(* Schneider Machine Expert - Basic project timer_options_behavior, file version 3.0.0.0 *)
(* ProjectInformations: Name=New project *)

HARDWARE
  Cpu 0: TM200CE40T
  EthernetConfiguration: NetworkName=M200, IpAllocationMode=FixedAddress, IpAddress=0.0.0.0, SubnetMask=0.0.0.0
  SerialLineConfiguration: Baud=Baud19200, Parity=ParityEven, DataBits=DataBits8, StopBits=StopBits1, PhysicalMedium=PhysicalMediumRs485, TransmissionMode=TransmissionModeModbusRtu, SlaveId=1, Addressing=SlaveAddressing
  MastTask: UsePeriodScanMode=false, PeriodScan=100
  FastTask: Period=255
  CpuBehavior: StartingMode=StartAsPreviousState, AutoSaveRamOnEeprom=true, WatchdogPeriod=250

SYMBOLS  (address, symbol, comment, settings)
  %M500     constant_false_500
  %M501     compiler_reused_M501_501
  %M502     compiler_reused_M502_502
  %M503     compiler_reused_M503_503
  %M504     compiler_reused_M504_504
  %M505     compiler_reused_M505_505
  %M506     compiler_reused_M506_506
  %M507     compiler_reused_M507_507
  %M508     compiler_reused_M508_508
  %M509     compiler_reused_M509_509
  %M510     output_5_image_510
  %M511     input_1_snapshot_511
  %M512     output_6_image_512
  %M513     input_0_snapshot_513
  %M514     output_7_image_514
  %M515     output_8_image_515
  %M516     output_9_image_516
  %M517     output_10_image_517
  %M518     output_11_image_518
  %M519     output_12_image_519
  %M520     output_13_image_520
  %M521     output_14_image_521
  %S13      SB_FIRSTRUN  "Indicates the first controller cycle in RUN mode"
  %MW4000   compiler_reused_MW4000_MW4000
  %TM0        [Preset=20, Base=OneSecond, IsRetentive=true]
  %TM1        [Type=TOF, Preset=20, Base=OneSecond, IsRetentive=true]
  %TM2        [Preset=20, Base=OneSecond, IsDynamicPreset=true]

POU Generated C++ - EXPERIMENTAL
  (* SectionNumber=1 *)

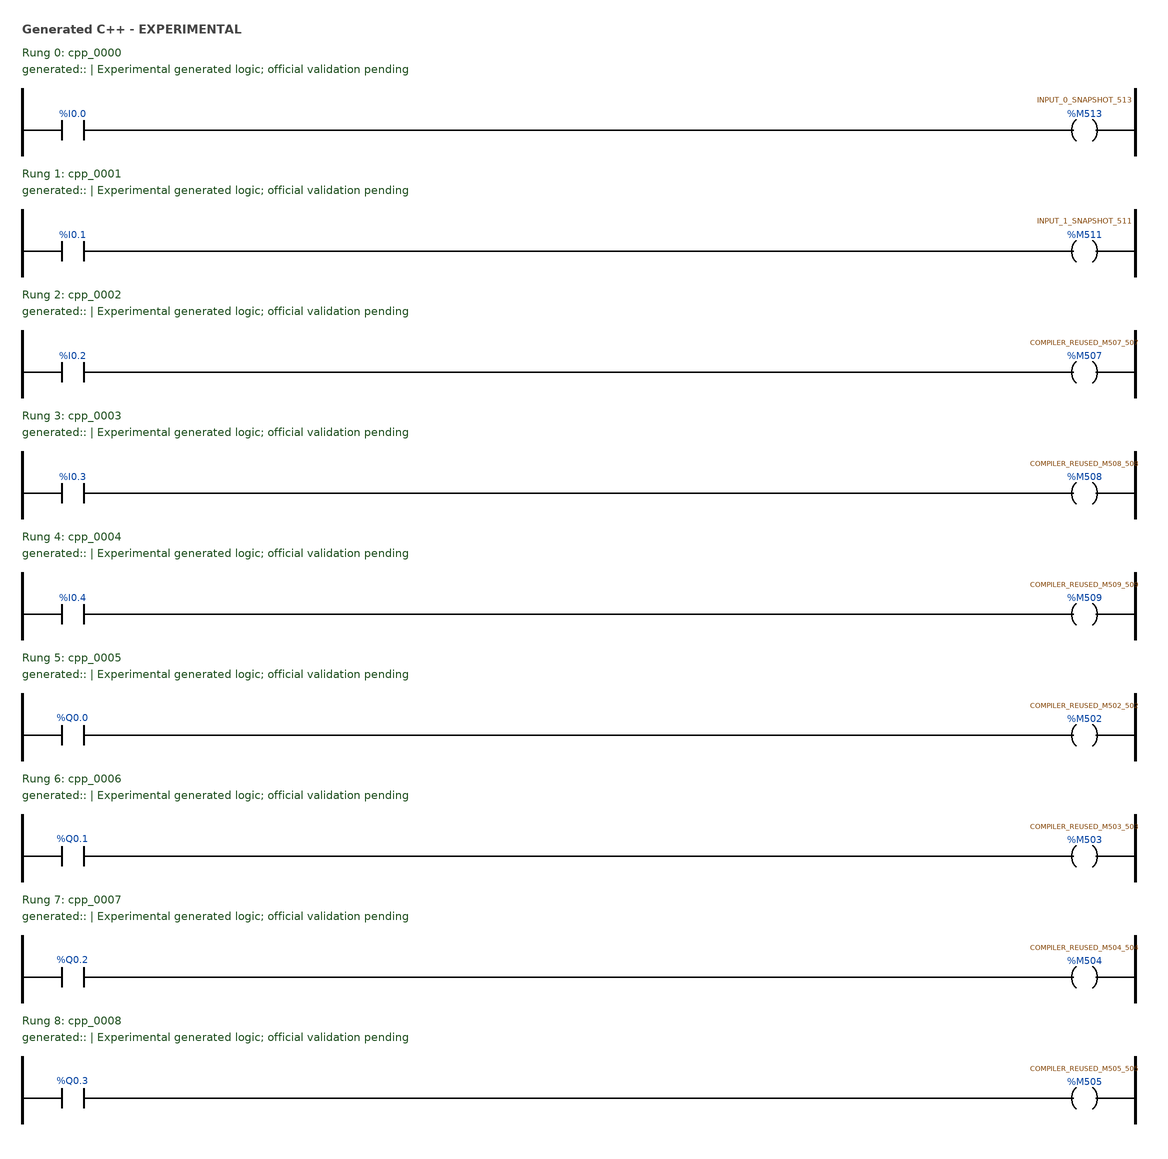

// Rung 0: cpp_0000
// generated:: | Experimental generated logic; official validation pending
  LD %I0.0
  ST %M513                (* input_0_snapshot_513 *)
  // as ST:
  //   input_0_snapshot_513 := %I0.0;

// Rung 1: cpp_0001
// generated:: | Experimental generated logic; official validation pending
  LD %I0.1
  ST %M511                (* input_1_snapshot_511 *)
  // as ST:
  //   input_1_snapshot_511 := %I0.1;

// Rung 2: cpp_0002
// generated:: | Experimental generated logic; official validation pending
  LD %I0.2
  ST %M507                (* compiler_reused_M507_507 *)
  // as ST:
  //   compiler_reused_M507_507 := %I0.2;

// Rung 3: cpp_0003
// generated:: | Experimental generated logic; official validation pending
  LD %I0.3
  ST %M508                (* compiler_reused_M508_508 *)
  // as ST:
  //   compiler_reused_M508_508 := %I0.3;

// Rung 4: cpp_0004
// generated:: | Experimental generated logic; official validation pending
  LD %I0.4
  ST %M509                (* compiler_reused_M509_509 *)
  // as ST:
  //   compiler_reused_M509_509 := %I0.4;

// Rung 5: cpp_0005
// generated:: | Experimental generated logic; official validation pending
  LD %Q0.0
  ST %M502                (* compiler_reused_M502_502 *)
  // as ST:
  //   compiler_reused_M502_502 := %Q0.0;

// Rung 6: cpp_0006
// generated:: | Experimental generated logic; official validation pending
  LD %Q0.1
  ST %M503                (* compiler_reused_M503_503 *)
  // as ST:
  //   compiler_reused_M503_503 := %Q0.1;

// Rung 7: cpp_0007
// generated:: | Experimental generated logic; official validation pending
  LD %Q0.2
  ST %M504                (* compiler_reused_M504_504 *)
  // as ST:
  //   compiler_reused_M504_504 := %Q0.2;

// Rung 8: cpp_0008
// generated:: | Experimental generated logic; official validation pending
  LD %Q0.3
  ST %M505                (* compiler_reused_M505_505 *)
  // as ST:
  //   compiler_reused_M505_505 := %Q0.3;

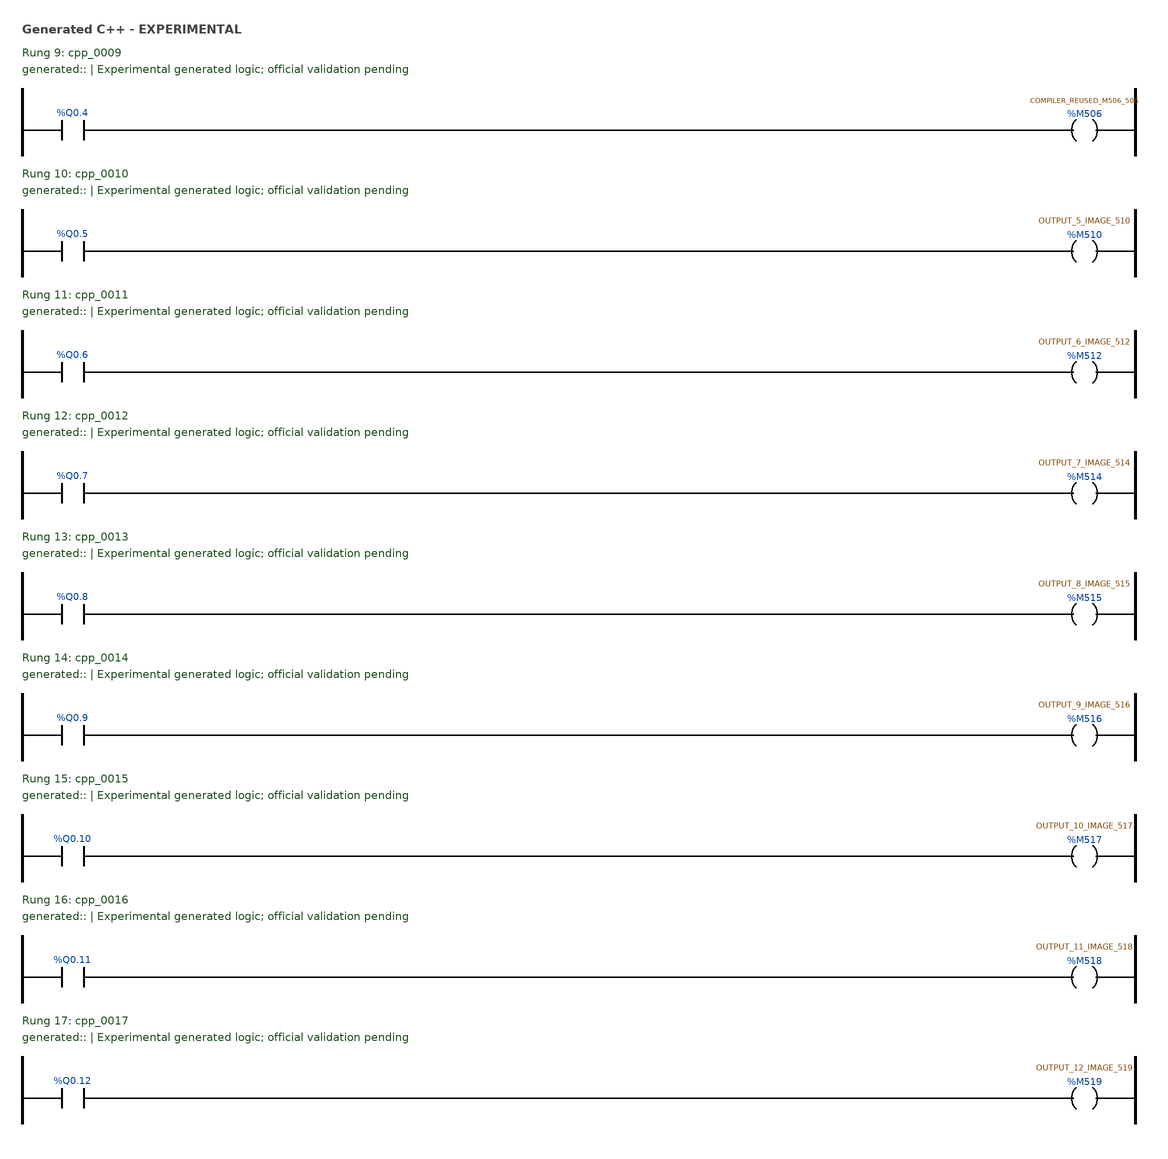

// Rung 9: cpp_0009
// generated:: | Experimental generated logic; official validation pending
  LD %Q0.4
  ST %M506                (* compiler_reused_M506_506 *)
  // as ST:
  //   compiler_reused_M506_506 := %Q0.4;

// Rung 10: cpp_0010
// generated:: | Experimental generated logic; official validation pending
  LD %Q0.5
  ST %M510                (* output_5_image_510 *)
  // as ST:
  //   output_5_image_510 := %Q0.5;

// Rung 11: cpp_0011
// generated:: | Experimental generated logic; official validation pending
  LD %Q0.6
  ST %M512                (* output_6_image_512 *)
  // as ST:
  //   output_6_image_512 := %Q0.6;

// Rung 12: cpp_0012
// generated:: | Experimental generated logic; official validation pending
  LD %Q0.7
  ST %M514                (* output_7_image_514 *)
  // as ST:
  //   output_7_image_514 := %Q0.7;

// Rung 13: cpp_0013
// generated:: | Experimental generated logic; official validation pending
  LD %Q0.8
  ST %M515                (* output_8_image_515 *)
  // as ST:
  //   output_8_image_515 := %Q0.8;

// Rung 14: cpp_0014
// generated:: | Experimental generated logic; official validation pending
  LD %Q0.9
  ST %M516                (* output_9_image_516 *)
  // as ST:
  //   output_9_image_516 := %Q0.9;

// Rung 15: cpp_0015
// generated:: | Experimental generated logic; official validation pending
  LD %Q0.10
  ST %M517                (* output_10_image_517 *)
  // as ST:
  //   output_10_image_517 := %Q0.10;

// Rung 16: cpp_0016
// generated:: | Experimental generated logic; official validation pending
  LD %Q0.11
  ST %M518                (* output_11_image_518 *)
  // as ST:
  //   output_11_image_518 := %Q0.11;

// Rung 17: cpp_0017
// generated:: | Experimental generated logic; official validation pending
  LD %Q0.12
  ST %M519                (* output_12_image_519 *)
  // as ST:
  //   output_12_image_519 := %Q0.12;

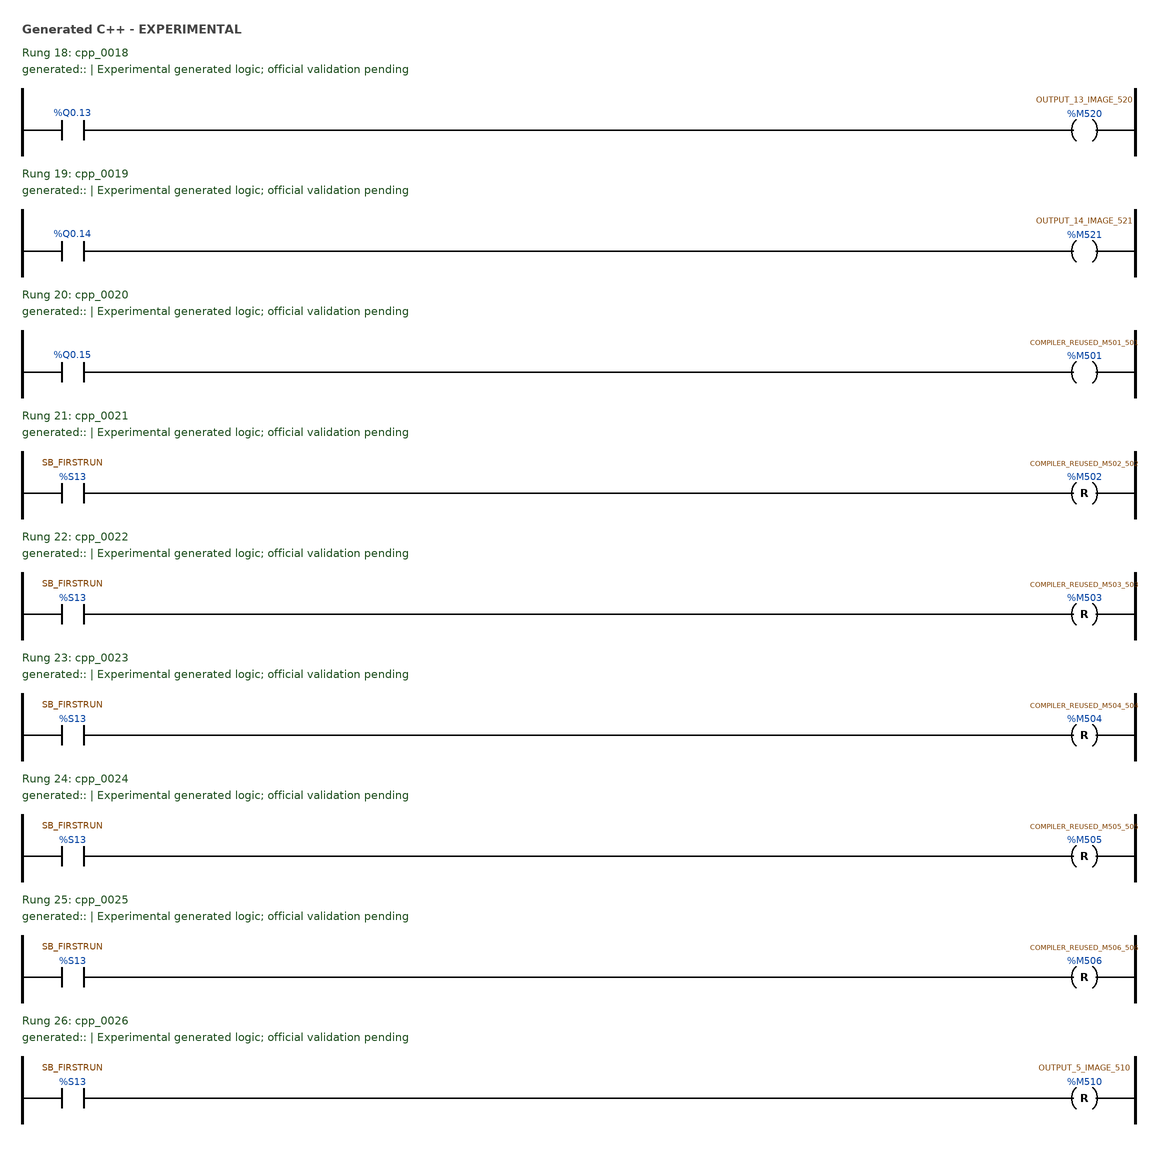

// Rung 18: cpp_0018
// generated:: | Experimental generated logic; official validation pending
  LD %Q0.13
  ST %M520                (* output_13_image_520 *)
  // as ST:
  //   output_13_image_520 := %Q0.13;

// Rung 19: cpp_0019
// generated:: | Experimental generated logic; official validation pending
  LD %Q0.14
  ST %M521                (* output_14_image_521 *)
  // as ST:
  //   output_14_image_521 := %Q0.14;

// Rung 20: cpp_0020
// generated:: | Experimental generated logic; official validation pending
  LD %Q0.15
  ST %M501                (* compiler_reused_M501_501 *)
  // as ST:
  //   compiler_reused_M501_501 := %Q0.15;

// Rung 21: cpp_0021
// generated:: | Experimental generated logic; official validation pending
  LD %S13                 (* SB_FIRSTRUN *)
  R %M502                 (* compiler_reused_M502_502 *)
  // as ST:
  //   IF SB_FIRSTRUN THEN compiler_reused_M502_502 := FALSE; END_IF;

// Rung 22: cpp_0022
// generated:: | Experimental generated logic; official validation pending
  LD %S13                 (* SB_FIRSTRUN *)
  R %M503                 (* compiler_reused_M503_503 *)
  // as ST:
  //   IF SB_FIRSTRUN THEN compiler_reused_M503_503 := FALSE; END_IF;

// Rung 23: cpp_0023
// generated:: | Experimental generated logic; official validation pending
  LD %S13                 (* SB_FIRSTRUN *)
  R %M504                 (* compiler_reused_M504_504 *)
  // as ST:
  //   IF SB_FIRSTRUN THEN compiler_reused_M504_504 := FALSE; END_IF;

// Rung 24: cpp_0024
// generated:: | Experimental generated logic; official validation pending
  LD %S13                 (* SB_FIRSTRUN *)
  R %M505                 (* compiler_reused_M505_505 *)
  // as ST:
  //   IF SB_FIRSTRUN THEN compiler_reused_M505_505 := FALSE; END_IF;

// Rung 25: cpp_0025
// generated:: | Experimental generated logic; official validation pending
  LD %S13                 (* SB_FIRSTRUN *)
  R %M506                 (* compiler_reused_M506_506 *)
  // as ST:
  //   IF SB_FIRSTRUN THEN compiler_reused_M506_506 := FALSE; END_IF;

// Rung 26: cpp_0026
// generated:: | Experimental generated logic; official validation pending
  LD %S13                 (* SB_FIRSTRUN *)
  R %M510                 (* output_5_image_510 *)
  // as ST:
  //   IF SB_FIRSTRUN THEN output_5_image_510 := FALSE; END_IF;

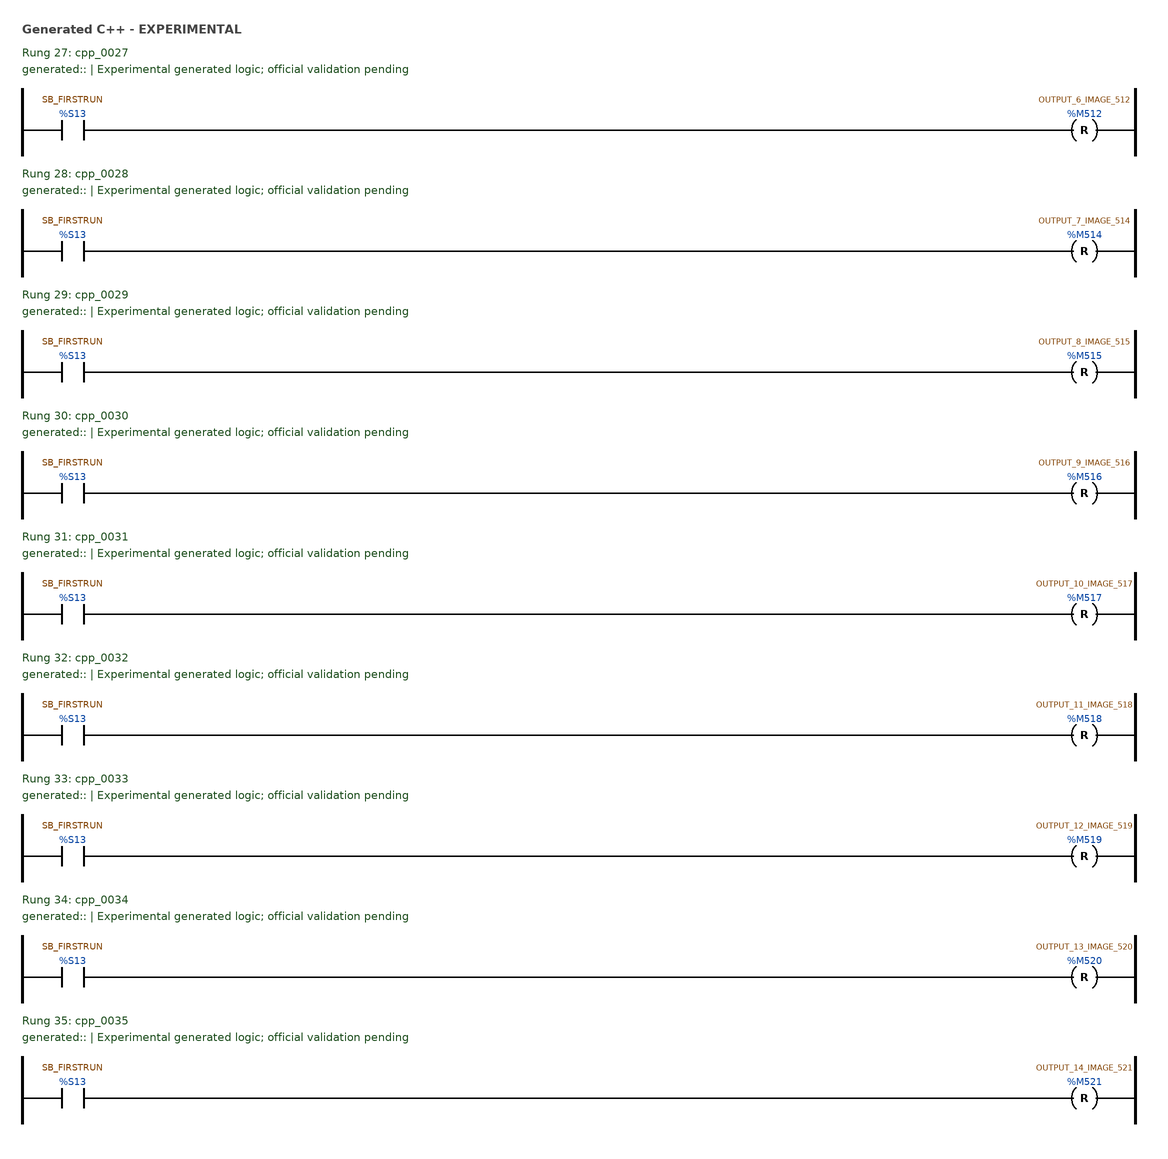

// Rung 27: cpp_0027
// generated:: | Experimental generated logic; official validation pending
  LD %S13                 (* SB_FIRSTRUN *)
  R %M512                 (* output_6_image_512 *)
  // as ST:
  //   IF SB_FIRSTRUN THEN output_6_image_512 := FALSE; END_IF;

// Rung 28: cpp_0028
// generated:: | Experimental generated logic; official validation pending
  LD %S13                 (* SB_FIRSTRUN *)
  R %M514                 (* output_7_image_514 *)
  // as ST:
  //   IF SB_FIRSTRUN THEN output_7_image_514 := FALSE; END_IF;

// Rung 29: cpp_0029
// generated:: | Experimental generated logic; official validation pending
  LD %S13                 (* SB_FIRSTRUN *)
  R %M515                 (* output_8_image_515 *)
  // as ST:
  //   IF SB_FIRSTRUN THEN output_8_image_515 := FALSE; END_IF;

// Rung 30: cpp_0030
// generated:: | Experimental generated logic; official validation pending
  LD %S13                 (* SB_FIRSTRUN *)
  R %M516                 (* output_9_image_516 *)
  // as ST:
  //   IF SB_FIRSTRUN THEN output_9_image_516 := FALSE; END_IF;

// Rung 31: cpp_0031
// generated:: | Experimental generated logic; official validation pending
  LD %S13                 (* SB_FIRSTRUN *)
  R %M517                 (* output_10_image_517 *)
  // as ST:
  //   IF SB_FIRSTRUN THEN output_10_image_517 := FALSE; END_IF;

// Rung 32: cpp_0032
// generated:: | Experimental generated logic; official validation pending
  LD %S13                 (* SB_FIRSTRUN *)
  R %M518                 (* output_11_image_518 *)
  // as ST:
  //   IF SB_FIRSTRUN THEN output_11_image_518 := FALSE; END_IF;

// Rung 33: cpp_0033
// generated:: | Experimental generated logic; official validation pending
  LD %S13                 (* SB_FIRSTRUN *)
  R %M519                 (* output_12_image_519 *)
  // as ST:
  //   IF SB_FIRSTRUN THEN output_12_image_519 := FALSE; END_IF;

// Rung 34: cpp_0034
// generated:: | Experimental generated logic; official validation pending
  LD %S13                 (* SB_FIRSTRUN *)
  R %M520                 (* output_13_image_520 *)
  // as ST:
  //   IF SB_FIRSTRUN THEN output_13_image_520 := FALSE; END_IF;

// Rung 35: cpp_0035
// generated:: | Experimental generated logic; official validation pending
  LD %S13                 (* SB_FIRSTRUN *)
  R %M521                 (* output_14_image_521 *)
  // as ST:
  //   IF SB_FIRSTRUN THEN output_14_image_521 := FALSE; END_IF;

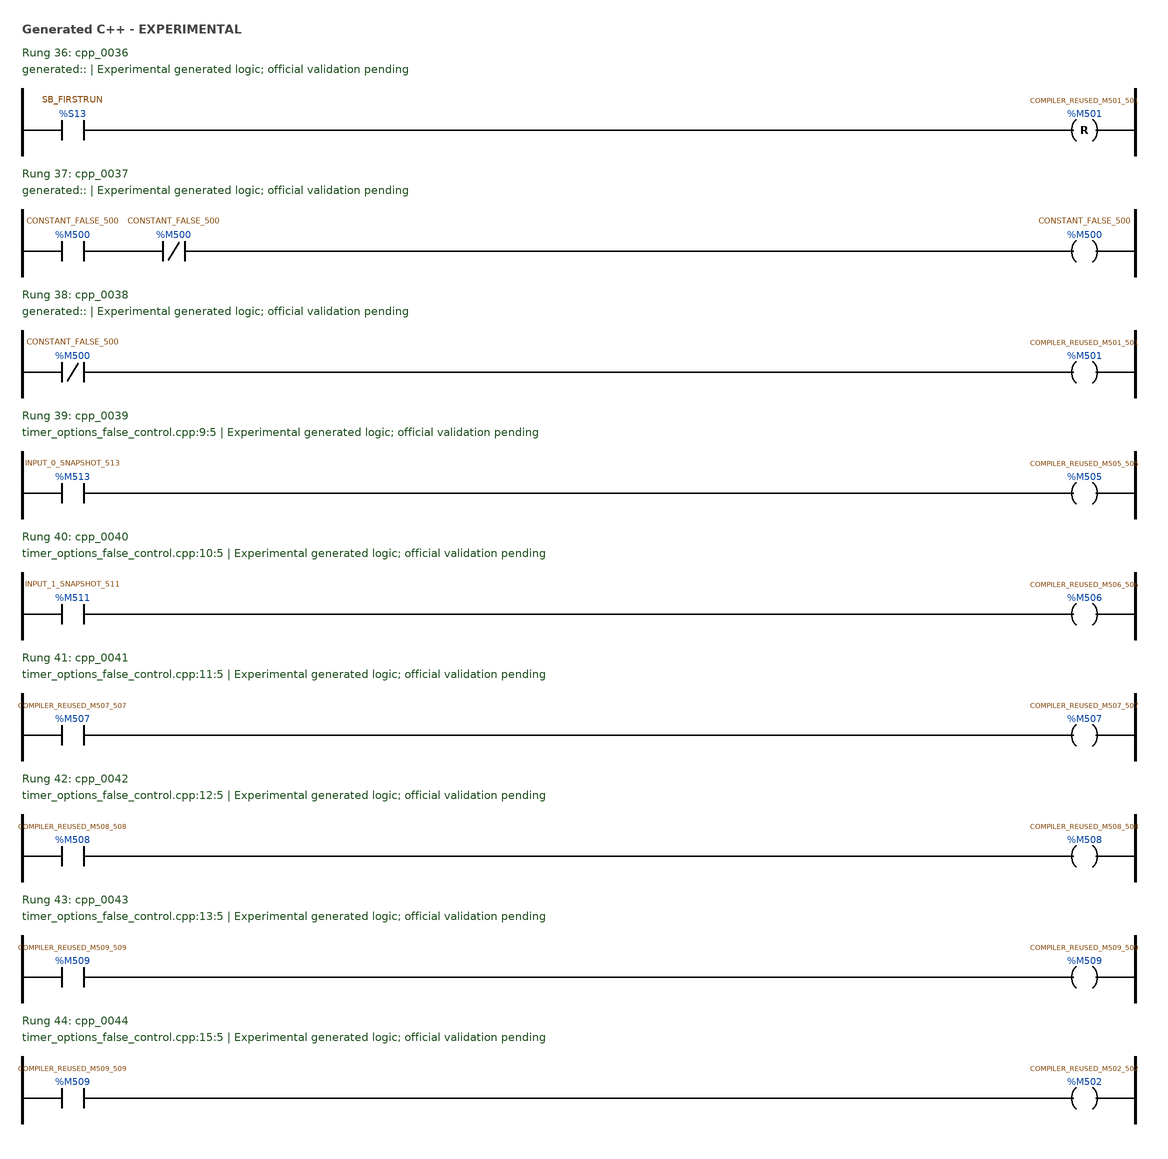

// Rung 36: cpp_0036
// generated:: | Experimental generated logic; official validation pending
  LD %S13                 (* SB_FIRSTRUN *)
  R %M501                 (* compiler_reused_M501_501 *)
  // as ST:
  //   IF SB_FIRSTRUN THEN compiler_reused_M501_501 := FALSE; END_IF;

// Rung 37: cpp_0037
// generated:: | Experimental generated logic; official validation pending
  LD %M500                (* constant_false_500 *)
  ANDN %M500              (* constant_false_500 *)
  ST %M500                (* constant_false_500 *)
  // as ST:
  //   constant_false_500 := constant_false_500 AND NOT constant_false_500;

// Rung 38: cpp_0038
// generated:: | Experimental generated logic; official validation pending
  LDN %M500               (* constant_false_500 *)
  ST %M501                (* compiler_reused_M501_501 *)
  // as ST:
  //   compiler_reused_M501_501 := NOT constant_false_500;

// Rung 39: cpp_0039
// timer_options_false_control.cpp:9:5 | Experimental generated logic; official validation pending
  LD %M513                (* input_0_snapshot_513 *)
  ST %M505                (* compiler_reused_M505_505 *)
  // as ST:
  //   compiler_reused_M505_505 := input_0_snapshot_513;

// Rung 40: cpp_0040
// timer_options_false_control.cpp:10:5 | Experimental generated logic; official validation pending
  LD %M511                (* input_1_snapshot_511 *)
  ST %M506                (* compiler_reused_M506_506 *)
  // as ST:
  //   compiler_reused_M506_506 := input_1_snapshot_511;

// Rung 41: cpp_0041
// timer_options_false_control.cpp:11:5 | Experimental generated logic; official validation pending
  LD %M507                (* compiler_reused_M507_507 *)
  ST %M507                (* compiler_reused_M507_507 *)
  // as ST:
  //   compiler_reused_M507_507 := compiler_reused_M507_507;

// Rung 42: cpp_0042
// timer_options_false_control.cpp:12:5 | Experimental generated logic; official validation pending
  LD %M508                (* compiler_reused_M508_508 *)
  ST %M508                (* compiler_reused_M508_508 *)
  // as ST:
  //   compiler_reused_M508_508 := compiler_reused_M508_508;

// Rung 43: cpp_0043
// timer_options_false_control.cpp:13:5 | Experimental generated logic; official validation pending
  LD %M509                (* compiler_reused_M509_509 *)
  ST %M509                (* compiler_reused_M509_509 *)
  // as ST:
  //   compiler_reused_M509_509 := compiler_reused_M509_509;

// Rung 44: cpp_0044
// timer_options_false_control.cpp:15:5 | Experimental generated logic; official validation pending
  LD %M509                (* compiler_reused_M509_509 *)
  ST %M502                (* compiler_reused_M502_502 *)
  // as ST:
  //   compiler_reused_M502_502 := compiler_reused_M509_509;

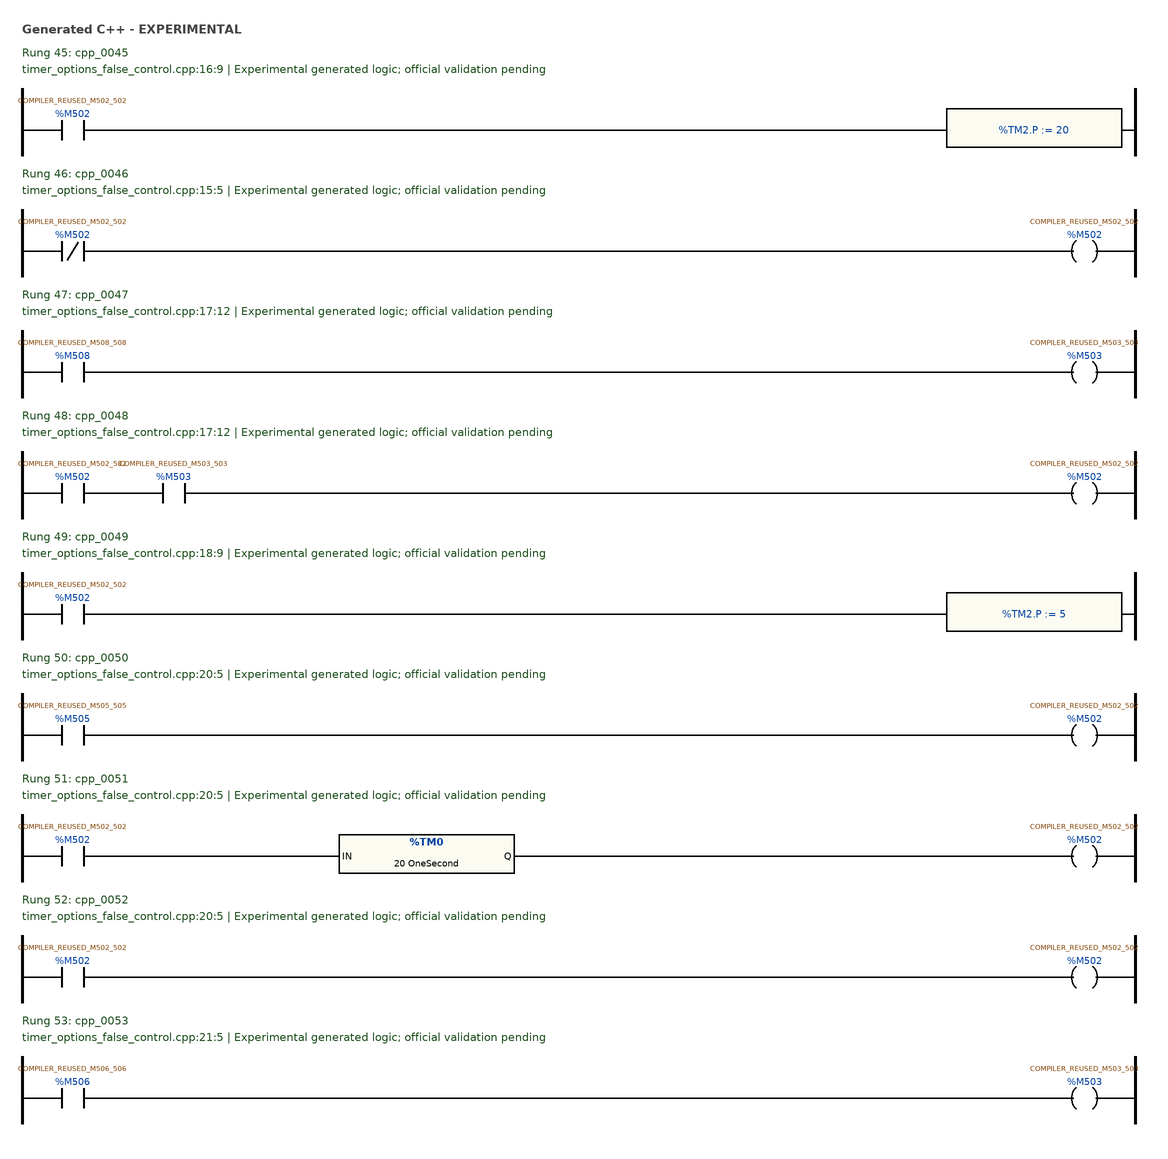

// Rung 45: cpp_0045
// timer_options_false_control.cpp:16:9 | Experimental generated logic; official validation pending
  LD %M502                (* compiler_reused_M502_502 *)
  [ %TM2.P := 20 ]
  // as ST:
  //   IF compiler_reused_M502_502 THEN %TM2.P := 20; END_IF;

// Rung 46: cpp_0046
// timer_options_false_control.cpp:15:5 | Experimental generated logic; official validation pending
  LDN %M502               (* compiler_reused_M502_502 *)
  ST %M502                (* compiler_reused_M502_502 *)
  // as ST:
  //   compiler_reused_M502_502 := NOT compiler_reused_M502_502;

// Rung 47: cpp_0047
// timer_options_false_control.cpp:17:12 | Experimental generated logic; official validation pending
  LD %M508                (* compiler_reused_M508_508 *)
  ST %M503                (* compiler_reused_M503_503 *)
  // as ST:
  //   compiler_reused_M503_503 := compiler_reused_M508_508;

// Rung 48: cpp_0048
// timer_options_false_control.cpp:17:12 | Experimental generated logic; official validation pending
  LD %M502                (* compiler_reused_M502_502 *)
  AND %M503               (* compiler_reused_M503_503 *)
  ST %M502                (* compiler_reused_M502_502 *)
  // as ST:
  //   compiler_reused_M502_502 := compiler_reused_M502_502 AND compiler_reused_M503_503;

// Rung 49: cpp_0049
// timer_options_false_control.cpp:18:9 | Experimental generated logic; official validation pending
  LD %M502                (* compiler_reused_M502_502 *)
  [ %TM2.P := 5 ]
  // as ST:
  //   IF compiler_reused_M502_502 THEN %TM2.P := 5; END_IF;

// Rung 50: cpp_0050
// timer_options_false_control.cpp:20:5 | Experimental generated logic; official validation pending
  LD %M505                (* compiler_reused_M505_505 *)
  ST %M502                (* compiler_reused_M502_502 *)
  // as ST:
  //   compiler_reused_M502_502 := compiler_reused_M505_505;

// Rung 51: cpp_0051
// timer_options_false_control.cpp:20:5 | Experimental generated logic; official validation pending
  BLK %TM0
  LD %M502                (* compiler_reused_M502_502 *)
  IN
  OUT_BLK
  LD Q
  ST %M502                (* compiler_reused_M502_502 *)
  END_BLK
  // as ST:
  //   %TM0(IN := compiler_reused_M502_502);
  //   compiler_reused_M502_502 := %TM0.Q;

// Rung 52: cpp_0052
// timer_options_false_control.cpp:20:5 | Experimental generated logic; official validation pending
  LD %M502                (* compiler_reused_M502_502 *)
  ST %M502                (* compiler_reused_M502_502 *)
  // as ST:
  //   compiler_reused_M502_502 := compiler_reused_M502_502;

// Rung 53: cpp_0053
// timer_options_false_control.cpp:21:5 | Experimental generated logic; official validation pending
  LD %M506                (* compiler_reused_M506_506 *)
  ST %M503                (* compiler_reused_M503_503 *)
  // as ST:
  //   compiler_reused_M503_503 := compiler_reused_M506_506;

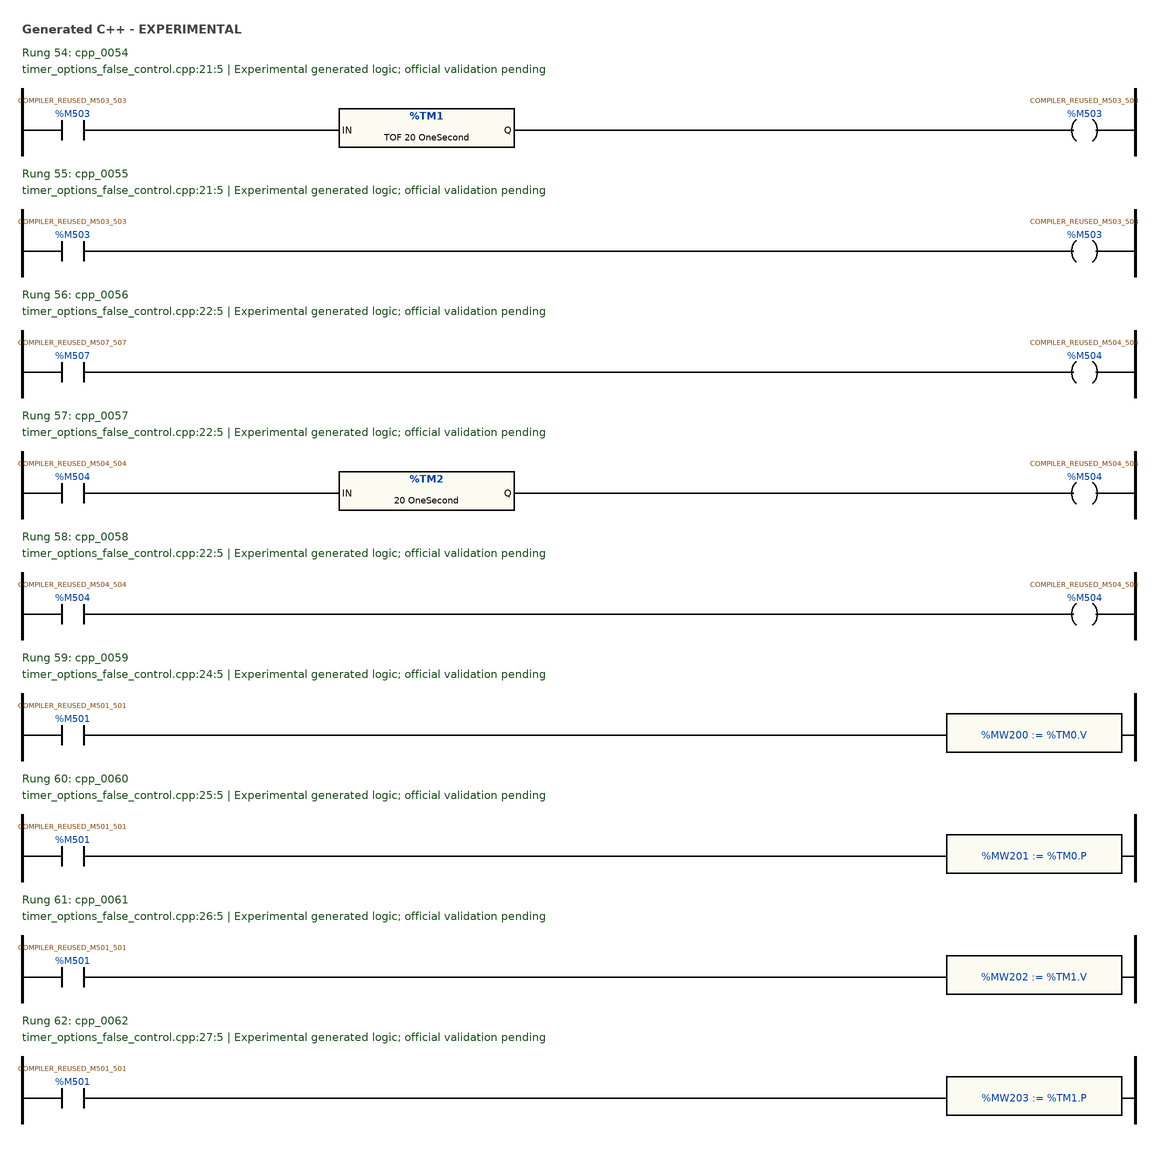

// Rung 54: cpp_0054
// timer_options_false_control.cpp:21:5 | Experimental generated logic; official validation pending
  BLK %TM1
  LD %M503                (* compiler_reused_M503_503 *)
  IN
  OUT_BLK
  LD Q
  ST %M503                (* compiler_reused_M503_503 *)
  END_BLK
  // as ST:
  //   %TM1(IN := compiler_reused_M503_503);
  //   compiler_reused_M503_503 := %TM1.Q;

// Rung 55: cpp_0055
// timer_options_false_control.cpp:21:5 | Experimental generated logic; official validation pending
  LD %M503                (* compiler_reused_M503_503 *)
  ST %M503                (* compiler_reused_M503_503 *)
  // as ST:
  //   compiler_reused_M503_503 := compiler_reused_M503_503;

// Rung 56: cpp_0056
// timer_options_false_control.cpp:22:5 | Experimental generated logic; official validation pending
  LD %M507                (* compiler_reused_M507_507 *)
  ST %M504                (* compiler_reused_M504_504 *)
  // as ST:
  //   compiler_reused_M504_504 := compiler_reused_M507_507;

// Rung 57: cpp_0057
// timer_options_false_control.cpp:22:5 | Experimental generated logic; official validation pending
  BLK %TM2
  LD %M504                (* compiler_reused_M504_504 *)
  IN
  OUT_BLK
  LD Q
  ST %M504                (* compiler_reused_M504_504 *)
  END_BLK
  // as ST:
  //   %TM2(IN := compiler_reused_M504_504);
  //   compiler_reused_M504_504 := %TM2.Q;

// Rung 58: cpp_0058
// timer_options_false_control.cpp:22:5 | Experimental generated logic; official validation pending
  LD %M504                (* compiler_reused_M504_504 *)
  ST %M504                (* compiler_reused_M504_504 *)
  // as ST:
  //   compiler_reused_M504_504 := compiler_reused_M504_504;

// Rung 59: cpp_0059
// timer_options_false_control.cpp:24:5 | Experimental generated logic; official validation pending
  LD %M501                (* compiler_reused_M501_501 *)
  [ %MW200 := %TM0.V ]
  // as ST:
  //   IF compiler_reused_M501_501 THEN %MW200 := %TM0.V; END_IF;

// Rung 60: cpp_0060
// timer_options_false_control.cpp:25:5 | Experimental generated logic; official validation pending
  LD %M501                (* compiler_reused_M501_501 *)
  [ %MW201 := %TM0.P ]
  // as ST:
  //   IF compiler_reused_M501_501 THEN %MW201 := %TM0.P; END_IF;

// Rung 61: cpp_0061
// timer_options_false_control.cpp:26:5 | Experimental generated logic; official validation pending
  LD %M501                (* compiler_reused_M501_501 *)
  [ %MW202 := %TM1.V ]
  // as ST:
  //   IF compiler_reused_M501_501 THEN %MW202 := %TM1.V; END_IF;

// Rung 62: cpp_0062
// timer_options_false_control.cpp:27:5 | Experimental generated logic; official validation pending
  LD %M501                (* compiler_reused_M501_501 *)
  [ %MW203 := %TM1.P ]
  // as ST:
  //   IF compiler_reused_M501_501 THEN %MW203 := %TM1.P; END_IF;

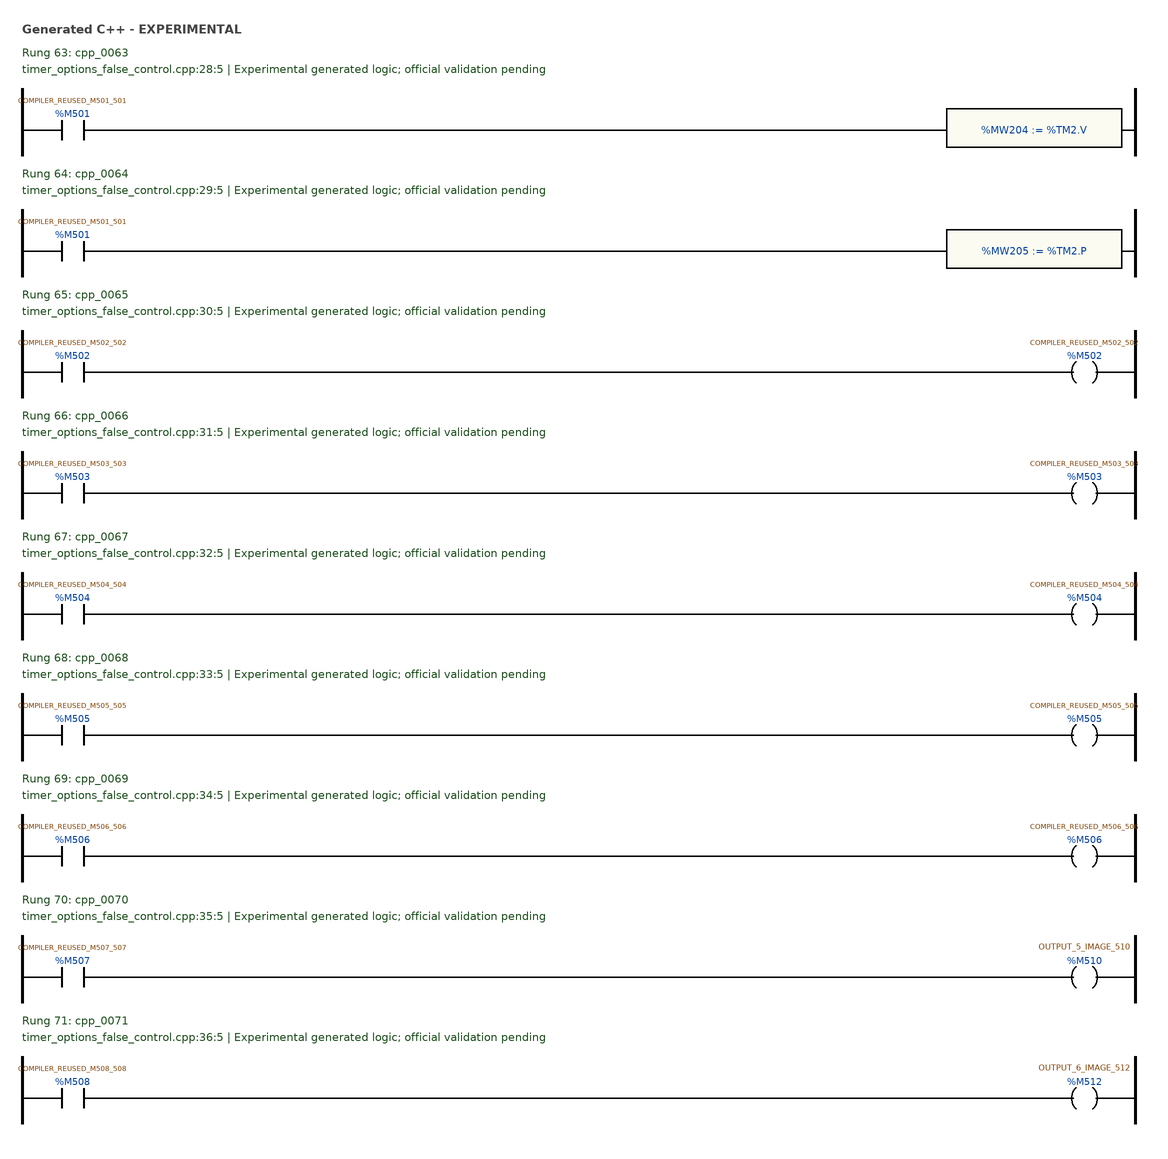

// Rung 63: cpp_0063
// timer_options_false_control.cpp:28:5 | Experimental generated logic; official validation pending
  LD %M501                (* compiler_reused_M501_501 *)
  [ %MW204 := %TM2.V ]
  // as ST:
  //   IF compiler_reused_M501_501 THEN %MW204 := %TM2.V; END_IF;

// Rung 64: cpp_0064
// timer_options_false_control.cpp:29:5 | Experimental generated logic; official validation pending
  LD %M501                (* compiler_reused_M501_501 *)
  [ %MW205 := %TM2.P ]
  // as ST:
  //   IF compiler_reused_M501_501 THEN %MW205 := %TM2.P; END_IF;

// Rung 65: cpp_0065
// timer_options_false_control.cpp:30:5 | Experimental generated logic; official validation pending
  LD %M502                (* compiler_reused_M502_502 *)
  ST %M502                (* compiler_reused_M502_502 *)
  // as ST:
  //   compiler_reused_M502_502 := compiler_reused_M502_502;

// Rung 66: cpp_0066
// timer_options_false_control.cpp:31:5 | Experimental generated logic; official validation pending
  LD %M503                (* compiler_reused_M503_503 *)
  ST %M503                (* compiler_reused_M503_503 *)
  // as ST:
  //   compiler_reused_M503_503 := compiler_reused_M503_503;

// Rung 67: cpp_0067
// timer_options_false_control.cpp:32:5 | Experimental generated logic; official validation pending
  LD %M504                (* compiler_reused_M504_504 *)
  ST %M504                (* compiler_reused_M504_504 *)
  // as ST:
  //   compiler_reused_M504_504 := compiler_reused_M504_504;

// Rung 68: cpp_0068
// timer_options_false_control.cpp:33:5 | Experimental generated logic; official validation pending
  LD %M505                (* compiler_reused_M505_505 *)
  ST %M505                (* compiler_reused_M505_505 *)
  // as ST:
  //   compiler_reused_M505_505 := compiler_reused_M505_505;

// Rung 69: cpp_0069
// timer_options_false_control.cpp:34:5 | Experimental generated logic; official validation pending
  LD %M506                (* compiler_reused_M506_506 *)
  ST %M506                (* compiler_reused_M506_506 *)
  // as ST:
  //   compiler_reused_M506_506 := compiler_reused_M506_506;

// Rung 70: cpp_0070
// timer_options_false_control.cpp:35:5 | Experimental generated logic; official validation pending
  LD %M507                (* compiler_reused_M507_507 *)
  ST %M510                (* output_5_image_510 *)
  // as ST:
  //   output_5_image_510 := compiler_reused_M507_507;

// Rung 71: cpp_0071
// timer_options_false_control.cpp:36:5 | Experimental generated logic; official validation pending
  LD %M508                (* compiler_reused_M508_508 *)
  ST %M512                (* output_6_image_512 *)
  // as ST:
  //   output_6_image_512 := compiler_reused_M508_508;

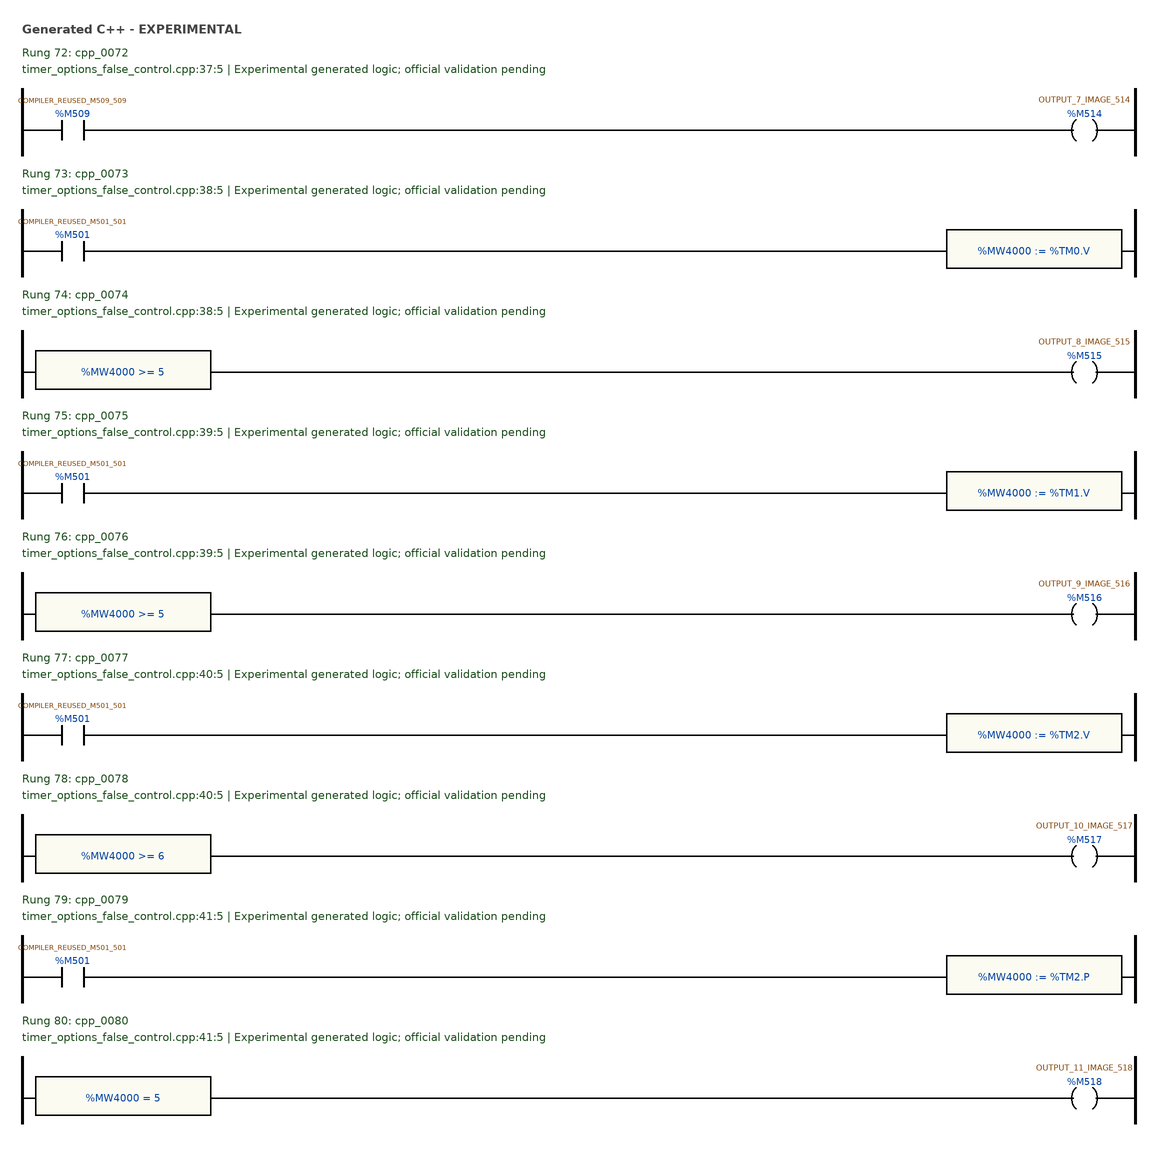

// Rung 72: cpp_0072
// timer_options_false_control.cpp:37:5 | Experimental generated logic; official validation pending
  LD %M509                (* compiler_reused_M509_509 *)
  ST %M514                (* output_7_image_514 *)
  // as ST:
  //   output_7_image_514 := compiler_reused_M509_509;

// Rung 73: cpp_0073
// timer_options_false_control.cpp:38:5 | Experimental generated logic; official validation pending
  LD %M501                (* compiler_reused_M501_501 *)
  [ %MW4000 := %TM0.V ]   (* compiler_reused_MW4000_MW4000 *)
  // as ST:
  //   IF compiler_reused_M501_501 THEN compiler_reused_MW4000_MW4000 := %TM0.V; END_IF;

// Rung 74: cpp_0074
// timer_options_false_control.cpp:38:5 | Experimental generated logic; official validation pending
  LD [ %MW4000 >= 5 ]     (* compiler_reused_MW4000_MW4000 *)
  ST %M515                (* output_8_image_515 *)
  // as ST:
  //   output_8_image_515 := compiler_reused_MW4000_MW4000 >= 5;

// Rung 75: cpp_0075
// timer_options_false_control.cpp:39:5 | Experimental generated logic; official validation pending
  LD %M501                (* compiler_reused_M501_501 *)
  [ %MW4000 := %TM1.V ]   (* compiler_reused_MW4000_MW4000 *)
  // as ST:
  //   IF compiler_reused_M501_501 THEN compiler_reused_MW4000_MW4000 := %TM1.V; END_IF;

// Rung 76: cpp_0076
// timer_options_false_control.cpp:39:5 | Experimental generated logic; official validation pending
  LD [ %MW4000 >= 5 ]     (* compiler_reused_MW4000_MW4000 *)
  ST %M516                (* output_9_image_516 *)
  // as ST:
  //   output_9_image_516 := compiler_reused_MW4000_MW4000 >= 5;

// Rung 77: cpp_0077
// timer_options_false_control.cpp:40:5 | Experimental generated logic; official validation pending
  LD %M501                (* compiler_reused_M501_501 *)
  [ %MW4000 := %TM2.V ]   (* compiler_reused_MW4000_MW4000 *)
  // as ST:
  //   IF compiler_reused_M501_501 THEN compiler_reused_MW4000_MW4000 := %TM2.V; END_IF;

// Rung 78: cpp_0078
// timer_options_false_control.cpp:40:5 | Experimental generated logic; official validation pending
  LD [ %MW4000 >= 6 ]     (* compiler_reused_MW4000_MW4000 *)
  ST %M517                (* output_10_image_517 *)
  // as ST:
  //   output_10_image_517 := compiler_reused_MW4000_MW4000 >= 6;

// Rung 79: cpp_0079
// timer_options_false_control.cpp:41:5 | Experimental generated logic; official validation pending
  LD %M501                (* compiler_reused_M501_501 *)
  [ %MW4000 := %TM2.P ]   (* compiler_reused_MW4000_MW4000 *)
  // as ST:
  //   IF compiler_reused_M501_501 THEN compiler_reused_MW4000_MW4000 := %TM2.P; END_IF;

// Rung 80: cpp_0080
// timer_options_false_control.cpp:41:5 | Experimental generated logic; official validation pending
  LD [ %MW4000 = 5 ]      (* compiler_reused_MW4000_MW4000 *)
  ST %M518                (* output_11_image_518 *)
  // as ST:
  //   output_11_image_518 := compiler_reused_MW4000_MW4000 = 5;

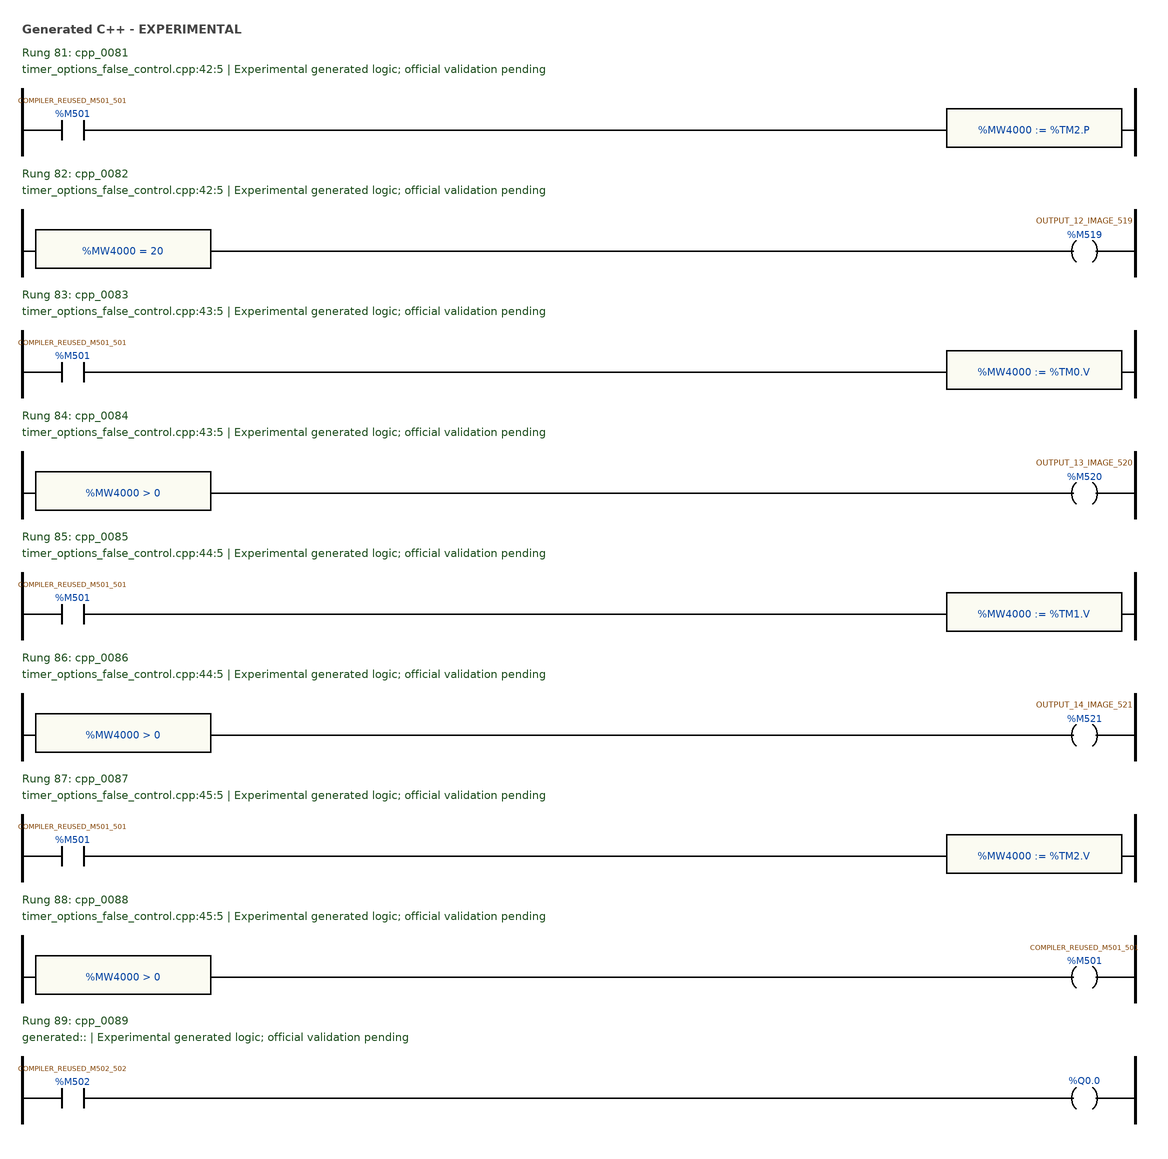

// Rung 81: cpp_0081
// timer_options_false_control.cpp:42:5 | Experimental generated logic; official validation pending
  LD %M501                (* compiler_reused_M501_501 *)
  [ %MW4000 := %TM2.P ]   (* compiler_reused_MW4000_MW4000 *)
  // as ST:
  //   IF compiler_reused_M501_501 THEN compiler_reused_MW4000_MW4000 := %TM2.P; END_IF;

// Rung 82: cpp_0082
// timer_options_false_control.cpp:42:5 | Experimental generated logic; official validation pending
  LD [ %MW4000 = 20 ]     (* compiler_reused_MW4000_MW4000 *)
  ST %M519                (* output_12_image_519 *)
  // as ST:
  //   output_12_image_519 := compiler_reused_MW4000_MW4000 = 20;

// Rung 83: cpp_0083
// timer_options_false_control.cpp:43:5 | Experimental generated logic; official validation pending
  LD %M501                (* compiler_reused_M501_501 *)
  [ %MW4000 := %TM0.V ]   (* compiler_reused_MW4000_MW4000 *)
  // as ST:
  //   IF compiler_reused_M501_501 THEN compiler_reused_MW4000_MW4000 := %TM0.V; END_IF;

// Rung 84: cpp_0084
// timer_options_false_control.cpp:43:5 | Experimental generated logic; official validation pending
  LD [ %MW4000 > 0 ]      (* compiler_reused_MW4000_MW4000 *)
  ST %M520                (* output_13_image_520 *)
  // as ST:
  //   output_13_image_520 := compiler_reused_MW4000_MW4000 > 0;

// Rung 85: cpp_0085
// timer_options_false_control.cpp:44:5 | Experimental generated logic; official validation pending
  LD %M501                (* compiler_reused_M501_501 *)
  [ %MW4000 := %TM1.V ]   (* compiler_reused_MW4000_MW4000 *)
  // as ST:
  //   IF compiler_reused_M501_501 THEN compiler_reused_MW4000_MW4000 := %TM1.V; END_IF;

// Rung 86: cpp_0086
// timer_options_false_control.cpp:44:5 | Experimental generated logic; official validation pending
  LD [ %MW4000 > 0 ]      (* compiler_reused_MW4000_MW4000 *)
  ST %M521                (* output_14_image_521 *)
  // as ST:
  //   output_14_image_521 := compiler_reused_MW4000_MW4000 > 0;

// Rung 87: cpp_0087
// timer_options_false_control.cpp:45:5 | Experimental generated logic; official validation pending
  LD %M501                (* compiler_reused_M501_501 *)
  [ %MW4000 := %TM2.V ]   (* compiler_reused_MW4000_MW4000 *)
  // as ST:
  //   IF compiler_reused_M501_501 THEN compiler_reused_MW4000_MW4000 := %TM2.V; END_IF;

// Rung 88: cpp_0088
// timer_options_false_control.cpp:45:5 | Experimental generated logic; official validation pending
  LD [ %MW4000 > 0 ]      (* compiler_reused_MW4000_MW4000 *)
  ST %M501                (* compiler_reused_M501_501 *)
  // as ST:
  //   compiler_reused_M501_501 := compiler_reused_MW4000_MW4000 > 0;

// Rung 89: cpp_0089
// generated:: | Experimental generated logic; official validation pending
  LD %M502                (* compiler_reused_M502_502 *)
  ST %Q0.0
  // as ST:
  //   %Q0.0 := compiler_reused_M502_502;

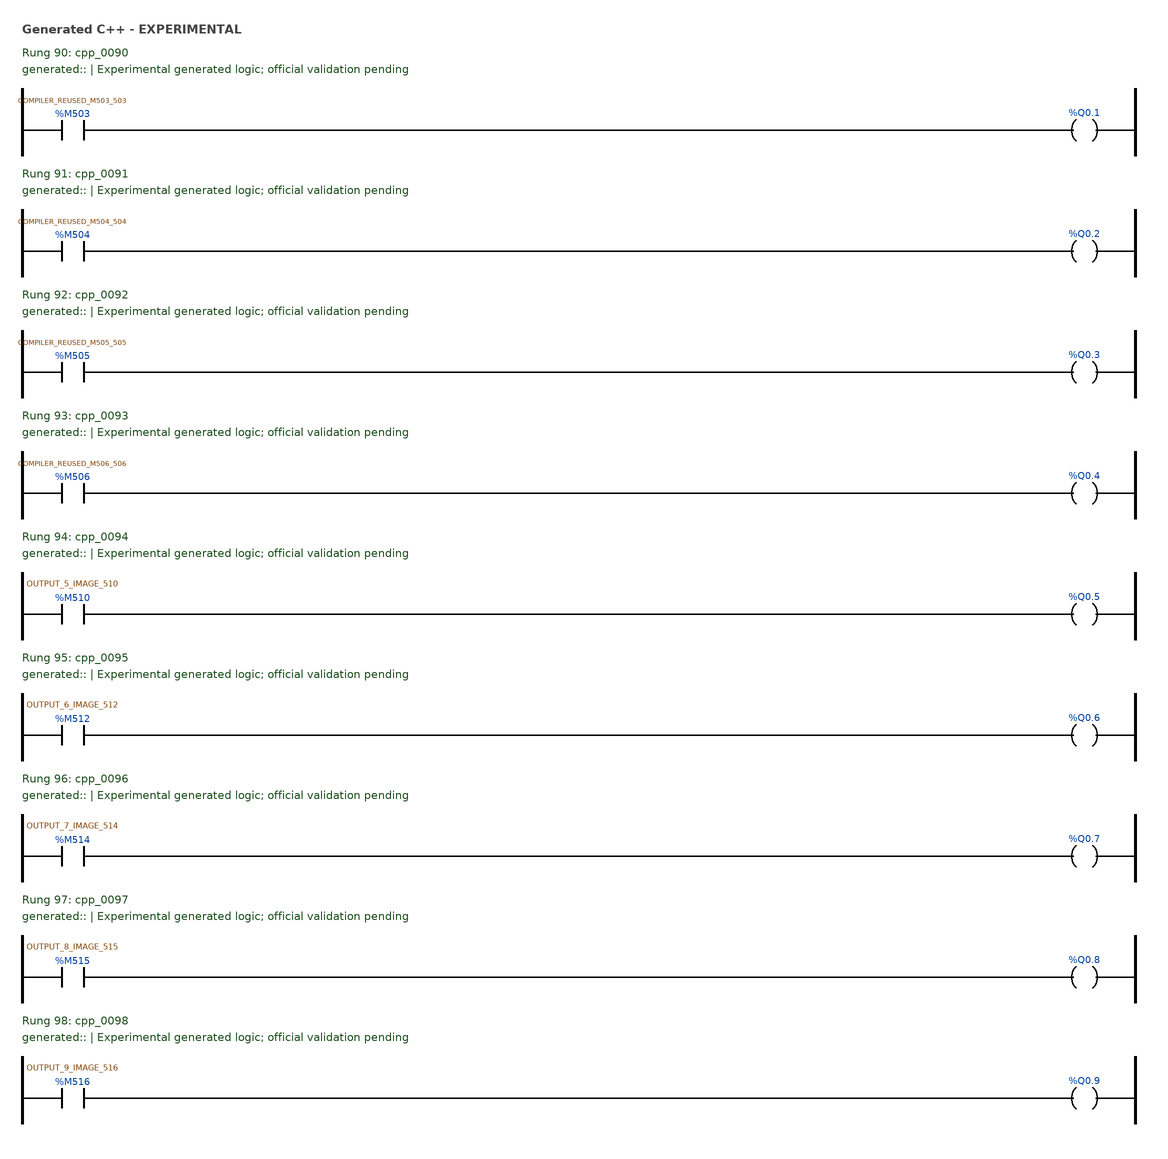

// Rung 90: cpp_0090
// generated:: | Experimental generated logic; official validation pending
  LD %M503                (* compiler_reused_M503_503 *)
  ST %Q0.1
  // as ST:
  //   %Q0.1 := compiler_reused_M503_503;

// Rung 91: cpp_0091
// generated:: | Experimental generated logic; official validation pending
  LD %M504                (* compiler_reused_M504_504 *)
  ST %Q0.2
  // as ST:
  //   %Q0.2 := compiler_reused_M504_504;

// Rung 92: cpp_0092
// generated:: | Experimental generated logic; official validation pending
  LD %M505                (* compiler_reused_M505_505 *)
  ST %Q0.3
  // as ST:
  //   %Q0.3 := compiler_reused_M505_505;

// Rung 93: cpp_0093
// generated:: | Experimental generated logic; official validation pending
  LD %M506                (* compiler_reused_M506_506 *)
  ST %Q0.4
  // as ST:
  //   %Q0.4 := compiler_reused_M506_506;

// Rung 94: cpp_0094
// generated:: | Experimental generated logic; official validation pending
  LD %M510                (* output_5_image_510 *)
  ST %Q0.5
  // as ST:
  //   %Q0.5 := output_5_image_510;

// Rung 95: cpp_0095
// generated:: | Experimental generated logic; official validation pending
  LD %M512                (* output_6_image_512 *)
  ST %Q0.6
  // as ST:
  //   %Q0.6 := output_6_image_512;

// Rung 96: cpp_0096
// generated:: | Experimental generated logic; official validation pending
  LD %M514                (* output_7_image_514 *)
  ST %Q0.7
  // as ST:
  //   %Q0.7 := output_7_image_514;

// Rung 97: cpp_0097
// generated:: | Experimental generated logic; official validation pending
  LD %M515                (* output_8_image_515 *)
  ST %Q0.8
  // as ST:
  //   %Q0.8 := output_8_image_515;

// Rung 98: cpp_0098
// generated:: | Experimental generated logic; official validation pending
  LD %M516                (* output_9_image_516 *)
  ST %Q0.9
  // as ST:
  //   %Q0.9 := output_9_image_516;

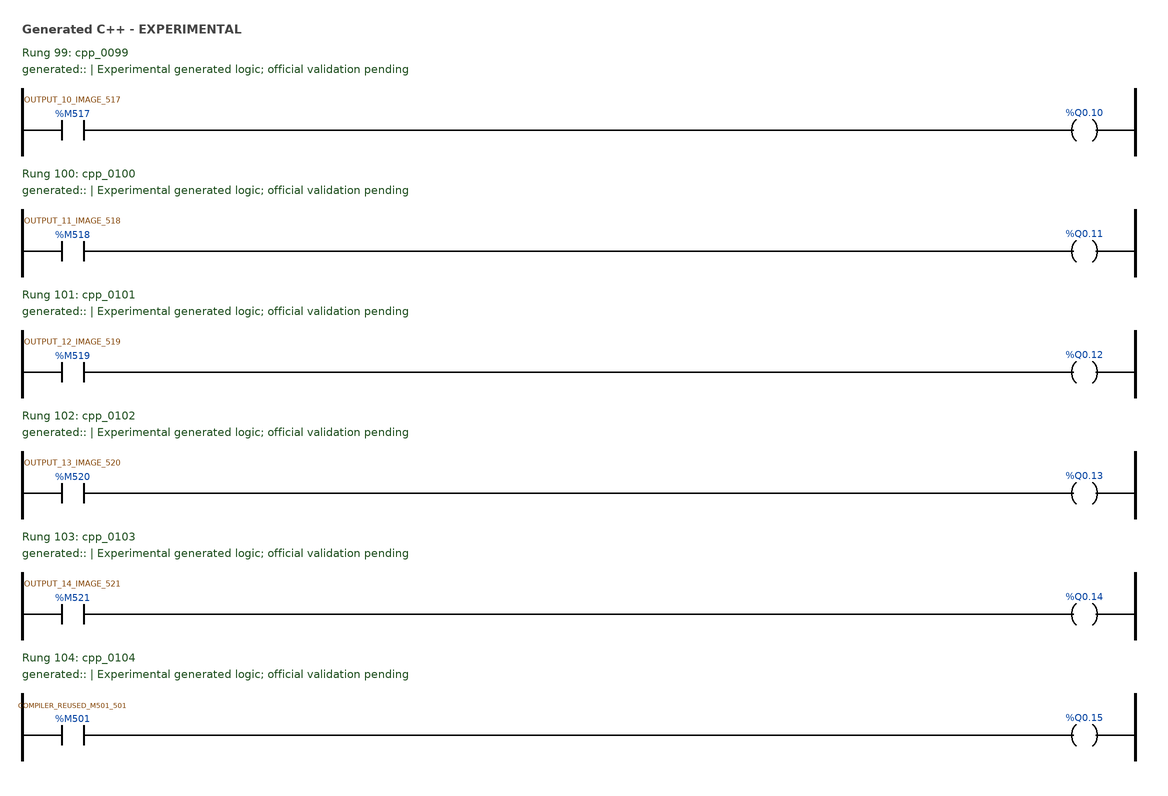

// Rung 99: cpp_0099
// generated:: | Experimental generated logic; official validation pending
  LD %M517                (* output_10_image_517 *)
  ST %Q0.10
  // as ST:
  //   %Q0.10 := output_10_image_517;

// Rung 100: cpp_0100
// generated:: | Experimental generated logic; official validation pending
  LD %M518                (* output_11_image_518 *)
  ST %Q0.11
  // as ST:
  //   %Q0.11 := output_11_image_518;

// Rung 101: cpp_0101
// generated:: | Experimental generated logic; official validation pending
  LD %M519                (* output_12_image_519 *)
  ST %Q0.12
  // as ST:
  //   %Q0.12 := output_12_image_519;

// Rung 102: cpp_0102
// generated:: | Experimental generated logic; official validation pending
  LD %M520                (* output_13_image_520 *)
  ST %Q0.13
  // as ST:
  //   %Q0.13 := output_13_image_520;

// Rung 103: cpp_0103
// generated:: | Experimental generated logic; official validation pending
  LD %M521                (* output_14_image_521 *)
  ST %Q0.14
  // as ST:
  //   %Q0.14 := output_14_image_521;

// Rung 104: cpp_0104
// generated:: | Experimental generated logic; official validation pending
  LD %M501                (* compiler_reused_M501_501 *)
  ST %Q0.15
  // as ST:
  //   %Q0.15 := compiler_reused_M501_501;
